(* IEC 61131-3 sources: volt/packages/volt-lsp-iec/test-corpus/awa-palletizer/Device/Plc Logic/Application/Library Manager/L_IE1P_ApplicationErrorsImplementation, 41 files *)

(* ---- L_IE1P_ERRORINFO.dut ---- *)
TYPE L_IE1P_ERRORINFO :
STRUCT
	XERROR : BOOL;
	WTEXTREFID : WORD;
	WERRORID : WORD;
	ESEVERITY : L_IE1P_SeverityLevel;
	EREACTION : L_IE1P_Reaction;
	EGROUP : L_IE1P_Group;
END_STRUCT
END_TYPE

(* ---- L_IE1P_ERRORINFORMATION.dut ---- *)
TYPE L_IE1P_ERRORINFORMATION :
STRUCT
	EERRORID : L_IE1P_Error;
	WCOMPID : WORD;
	ESEVERITY : L_IE1P_SeverityLevel;
	PSINSTANCENAME : POINTER TO STRING;
	INSTANCEID : DWORD := 0;
	TTIMESTAMP : TIME;
	TRESETTIMESTAMP : TIME;
	XCYCLIC : BOOL;
	DWEXTENDEDERRORINFO : DWORD;
	XEXTERNALERROR : BOOL;
	XCLEARERRORNEEDED : BOOL;
END_STRUCT
END_TYPE

(* ---- L_IE1P_INSTANCEIDS.dut ---- *)
TYPE L_IE1P_INSTANCEIDS :
STRUCT
	EXTINSTANCEID : DWORD;
	ADDINSTANCID1 : DWORD;
	ADDINSTANCID2 : DWORD;
	ADDINSTANCID3 : DWORD;
	ADDINSTANCID4 : DWORD;
END_STRUCT
END_TYPE

(* ---- L_IE1P_PARAMETERITEMMID.dut ---- *)
TYPE L_IE1P_PARAMETERITEMMID :
STRUCT
	SIZE : BYTE;
	ETYPE : INT;
	VALUE : L_IE1P_ParaValueMid;
END_STRUCT
END_TYPE

(* ---- L_IE1P_PARAVALUEMID.dut ---- *)
TYPE L_IE1P_PARAVALUEMID :
UNION
	DWVALUE : DWORD;
	DIVALUE : DINT;
	LRVALUE : REAL;
	SVALUE : STRING;
END_UNION
END_TYPE

(* ---- L_IE1P_PLACEHOLDERTYPE.dut ---- *)
TYPE L_IE1P_PLACEHOLDERTYPE :
(
	VTNONE := 0,
	VTDINT := 4,
	VTDWORD := 7,
	VTSTRING := 9
);
END_TYPE

(* ---- L_IE1P_PLACEHOLDERVALUE.dut ---- *)
TYPE L_IE1P_PLACEHOLDERVALUE :
UNION
	DIVALUE : DINT;
	DWVALUE : DWORD;
	RVALUE : REAL;
	LRVALUE : LREAL;
	SVALUE : STRING(50);
END_UNION
END_TYPE

(* ---- L_IE1P_PLACEHOLDERVARIABLE.dut ---- *)
TYPE L_IE1P_PLACEHOLDERVARIABLE :
STRUCT
	VARTYPE : L_IE1P_PlaceHolderType;
	VALUE : L_IE1P_PlaceholderValue;
END_STRUCT
END_TYPE

(* ---- L_IE1P_INTERNAL.gvl ---- *)
VAR_GLOBAL
	DEVICEEVENTMONITOR : L_IE1P_DeviceEventMonitor;
END_VAR

(* ---- L_IE1P_IATTRIBUTES.itf ---- *)
INTERFACE L_IE1P_IATTRIBUTES
END_INTERFACE

METHOD GET1STATTRIBUTE : DINT
END_METHOD

METHOD GET2NDATTRIBUTE : LREAL
END_METHOD

METHOD GET3RDATTRIBUTE : STRING(20)
END_METHOD

(* ---- L_IE1P_ITEXTPLACEHOLDER.itf ---- *)
INTERFACE L_IE1P_ITEXTPLACEHOLDER
END_INTERFACE

METHOD GETPLACEHOLDERDATA : L_IE1P_PlaceHolderType
VAR_INPUT
	INDEX : WORD;
END_VAR
VAR_OUTPUT
	PDATA : POINTER TO BYTE;
END_VAR
END_METHOD

(* ---- GETBOOLEANPROPERTY.pou ---- *)
FUNCTION GETBOOLEANPROPERTY : BOOL
VAR_INPUT
	STKEY : WSTRING;
END_VAR
END_FUNCTION

(* ---- GETCOMPANY.pou ---- *)
FUNCTION GETCOMPANY : WSTRING
END_FUNCTION

(* ---- GETNUMBERPROPERTY.pou ---- *)
FUNCTION GETNUMBERPROPERTY : DINT
VAR_INPUT
	STKEY : WSTRING;
END_VAR
END_FUNCTION

(* ---- GETTEXTPROPERTY.pou ---- *)
FUNCTION GETTEXTPROPERTY : WSTRING
VAR_INPUT
	STKEY : WSTRING;
END_VAR
END_FUNCTION

(* ---- GETTEXTPROPERTY2.pou ---- *)
FUNCTION GETTEXTPROPERTY2 : POINTER TO WSTRING
VAR_INPUT
	STKEY : WSTRING;
END_VAR
END_FUNCTION

(* ---- GETTITLE.pou ---- *)
FUNCTION GETTITLE : WSTRING
END_FUNCTION

(* ---- GETVERSION.pou ---- *)
FUNCTION GETVERSION : VERSION
END_FUNCTION

(* ---- GETVERSIONPROPERTY.pou ---- *)
FUNCTION GETVERSIONPROPERTY : VERSION
VAR_INPUT
	STKEY : WSTRING;
END_VAR
END_FUNCTION

(* ---- L_IE1P_GETHIGHESTREACTION.pou ---- *)
FUNCTION L_IE1P_GETHIGHESTREACTION : BOOL
VAR_INPUT
	EREACTION1 : L_IE1P_Reaction;
	MODULEHANDLER1 : POINTER TO BYTE;
	EREACTION2 : L_IE1P_Reaction;
	MODULEHANDLER2 : POINTER TO BYTE;
END_VAR
VAR_OUTPUT
	EREACTION : L_IE1P_Reaction;
	MODULEHANDLER : POINTER TO BYTE;
END_VAR
END_FUNCTION

(* ---- L_IE1P_GETHIGHESTSEVERITYANDREACTION.pou ---- *)
FUNCTION L_IE1P_GETHIGHESTSEVERITYANDREACTION : BOOL
VAR_INPUT
	ESEVERITY1 : L_IE1P_SeverityLevel;
	EREACTION1 : L_IE1P_Reaction;
	MODULEHANDLER1 : POINTER TO BYTE;
	ESEVERITY2 : L_IE1P_SeverityLevel;
	EREACTION2 : L_IE1P_Reaction;
	MODULEHANDLER2 : POINTER TO BYTE;
END_VAR
VAR_OUTPUT
	ESEVERITY : L_IE1P_SeverityLevel;
	EREACTION : L_IE1P_Reaction;
	MODULEHANDLER : POINTER TO BYTE;
END_VAR
END_FUNCTION

(* ---- L_IE1P_READERRORDATAFROMCOMPONENTLIST.pou ---- *)
FUNCTION L_IE1P_READERRORDATAFROMCOMPONENTLIST : BOOL
VAR_INPUT
	MODULEHANDLE : UDINT;
	PDATA : POINTER TO L_IE1P_ReadErrorData;
END_VAR
VAR_OUTPUT
	SEVERITY : L_IE1P_SeverityLevel;
	ERRORCODE : DWORD := 0;
END_VAR
VAR_IN_OUT
	DWCOMPIDX : DWORD;
END_VAR
END_FUNCTION

(* ---- GLOBALTEXTLIST.pou ---- *)
FUNCTION_BLOCK GLOBALTEXTLIST
VAR
	M_TEXTLISTFILE : STRING(255);
	_STNAMESPACE : STRING;
END_VAR
END_FUNCTION_BLOCK

(* ---- L_IE1P_ATTRIBUTES.pou ---- *)
FUNCTION_BLOCK L_IE1P_ATTRIBUTES
VAR_INPUT
	DIATTRIBUTE1 : DINT;
	LRATTRIBUTE2 : LREAL;
	SATTRIBUTE3 : STRING(20);
END_VAR
END_FUNCTION_BLOCK

METHOD GET1STATTRIBUTE : DINT
END_METHOD

METHOD GET2NDATTRIBUTE : LREAL
END_METHOD

METHOD GET3RDATTRIBUTE : STRING(20)
END_METHOD

(* ---- L_IE1P_DEVICEEVENTMONITOR.pou ---- *)
FUNCTION_BLOCK L_IE1P_DEVICEEVENTMONITOR
VAR
	ITFCALLBACK : CmpEventMgr.ICmpEventCallback;
	HEVENTACTUALERROR : SysTypes.RTS_IEC_HANDLE := SysTypes.RTS_INVALID_HANDLE;
	HINTERFACEACTUALERROR : SysTypes.RTS_IEC_HANDLE := SysTypes.RTS_INVALID_HANDLE;
	DWERRORUPDATED : DWORD := 0;
	AEACTSEVERITY : ARRAY [1..2] OF L_IE1P_SeverityLevel;
	ADWACTERRORCODE : ARRAY [1..2] OF DWORD;
	USIACTIVEERRORINFO : USINT;
END_VAR
END_FUNCTION_BLOCK

METHOD READACTUALERRORCODE
VAR_OUTPUT
	ESEVERITY : USINT;
	EREACTION : WORD;
	DWERRORCODE : DWORD;
END_VAR
END_METHOD

METHOD EVENTCALLBACK : UDINT
VAR_INPUT
	PEVENTPARAM : POINTER TO EventParam;
END_VAR
END_METHOD

METHOD REGISTEREVENT
VAR_INPUT
	XONLYCALLBACKFUNCTION : BOOL;
END_VAR
END_METHOD

METHOD UNREGISTEREVENT
VAR_INPUT
	XONLYCALLBACKFUNCTION : BOOL;
END_VAR
END_METHOD

METHOD FB_REINIT : BOOL
END_METHOD

METHOD FB_EXIT : BOOL
VAR_INPUT
	BINCOPYCODE : BOOL;
END_VAR
END_METHOD

METHOD FB_INIT : BOOL
VAR_INPUT
	BINITRETAINS : BOOL;
	BINCOPYCODE : BOOL;
END_VAR
END_METHOD

(* ---- L_IE1P_EMPTYERRORHANDLER.pou ---- *)
FUNCTION_BLOCK L_IE1P_EMPTYERRORHANDLER
END_FUNCTION_BLOCK

METHOD ITFCHECKERRORRESETOCCURED : BOOL
VAR_IN_OUT
	RESETTIME : SYSTIME;
END_VAR
END_METHOD

METHOD ITFCLEARERROR : DWORD
VAR_INPUT
	ESEVERITY : L_IE1P_SeverityLevel;
	WERRORID : WORD;
	WCOMPID : WORD;
	DWINSTANCEID : DWORD := 0;
END_VAR
END_METHOD

METHOD ITFCLEARREACTION
VAR_INPUT
	EREACTION : L_IE1P_Reaction;
	DICLEARCOUNT : DINT;
	DWINSTANCEID : DWORD;
END_VAR
END_METHOD

METHOD ITFGETACTUALERRORCODE : DWORD
VAR_OUTPUT
	ESEVERITY : WORD;
END_VAR
END_METHOD

METHOD ITFREGISTERERRORINSTANCE : DWORD
END_METHOD

METHOD ITFRESETACTIVE : BOOL
END_METHOD

METHOD ITFRESETERROR : DWORD
VAR_INPUT
	ERRORHANDLE : RTS_IEC_HANDLE := 0;
END_VAR
END_METHOD

METHOD ITFRESETERRORREACTION
VAR_INPUT
	DWINSTANCEID : DWORD := 0;
END_VAR
END_METHOD

METHOD ITFSETERROR : DWORD
VAR_INPUT
	ESEVERITY : L_IE1P_SeverityLevel;
	WERRORID : WORD;
	WCOMPID : WORD;
	DWINSTANCEID : DWORD := 0;
	EREACTION : L_IE1P_Reaction;
END_VAR
END_METHOD

(* ---- L_IE1P_ERRORHANDLER.pou ---- *)
FUNCTION_BLOCK L_IE1P_ERRORHANDLER
VAR_INPUT
	ADDERRORHANDLER1 : L_IE1P_IErrorHandler;
	ADDERRORHANDLER2 : L_IE1P_IErrorHandler;
	ADDERRORHANDLER3 : L_IE1P_IErrorHandler;
	ADDERRORHANDLER4 : L_IE1P_IErrorHandler;
END_VAR
VAR_OUTPUT
	XWARNINGACTIVE : BOOL;
	XWARNINGLOCKACTIVE : BOOL;
	XFAULTQSPAPPLACTIVE : BOOL;
	XFAULTQSPACTIVE : BOOL;
	XFAULTQSPCINHACTIVE : BOOL;
	XFAULTACTIVE : BOOL;
END_VAR
VAR
	ERRORMANAGER : L_IE1P_ErrorManager;
	ADDERRORHANDLERINSTANCEIDS : ARRAY [1..MaxInstanceIDs] OF L_IE1P_InstanceIDs;
	ERRORRESETOCCUREDTIME : SysTime;
	C_STRUNDEFERROR : STRING := 'undefined';
	MAXINSTANCEIDS : WORD := 15;
END_VAR
END_FUNCTION_BLOCK

METHOD CHECKHIGHESTSEVERITY
VAR_INPUT
	ESEVERITYNEW : WORD;
	DWERRORCODENEW : DWORD;
END_VAR
VAR_IN_OUT
	ESEVERITYACT : WORD;
	DWERRORCODEACT : DWORD;
END_VAR
END_METHOD

METHOD FINDADDINSTANCEID : DWORD
VAR_INPUT
	DWEXTINSTANCEID : DWORD;
	DWNUMBER : DWORD;
END_VAR
END_METHOD

METHOD FB_INIT : BOOL
VAR_INPUT
	BINITRETAINS : BOOL;
	BINCOPYCODE : BOOL;
END_VAR
END_METHOD

METHOD ITFCHECKERRORRESETOCCURED : BOOL
VAR_IN_OUT
	RESETTIME : SYSTIME;
END_VAR
END_METHOD

METHOD ITFCLEARERROR : DWORD
VAR_INPUT
	ESEVERITY : L_IE1P_SeverityLevel;
	WERRORID : WORD;
	WCOMPID : WORD;
	DWINSTANCEID : DWORD := 0;
END_VAR
END_METHOD

METHOD ITFCLEARREACTION
VAR_INPUT
	EREACTION : L_IE1P_Reaction;
	DICLEARCOUNT : DINT;
	DWINSTANCEID : DWORD;
END_VAR
END_METHOD

METHOD ITFGETACTUALERRORCODE : DWORD
VAR_OUTPUT
	ESEVERITY : WORD;
END_VAR
END_METHOD

METHOD ITFREGISTERERRORINSTANCE : DWORD
END_METHOD

METHOD ITFRESETACTIVE : BOOL
END_METHOD

METHOD ITFRESETERROR : DWORD
VAR_INPUT
	ERRORHANDLE : RTS_IEC_HANDLE := 0;
END_VAR
END_METHOD

METHOD ITFRESETERRORREACTION
VAR_INPUT
	DWINSTANCEID : DWORD := 0;
END_VAR
END_METHOD

METHOD ITFSETERROR : DWORD
VAR_INPUT
	ESEVERITY : L_IE1P_SeverityLevel;
	WERRORID : WORD;
	WCOMPID : WORD;
	DWINSTANCEID : DWORD := 0;
	EREACTION : L_IE1P_Reaction;
END_VAR
END_METHOD

(* ---- L_IE1P_ERRORMANAGER.pou ---- *)
FUNCTION_BLOCK L_IE1P_ERRORMANAGER
VAR_INPUT
	XUSEADDLOGIPC : BOOL := TRUE;
	DWTASKYCLE_US : DWORD := 1000;
	XIGNOREFAULT_LOG : BOOL := TRUE;
	XNOLOGBOOKENTRY : BOOL := FALSE;
END_VAR
VAR
	EACTIVEERRORID : REFERENCE TO L_IE1P_Error;
	EACTIVESEVERITY : REFERENCE TO L_IE1P_SeverityLevel;
	XERROR : REFERENCE TO BOOL;
	XWARNING : REFERENCE TO BOOL;
	PSERRORINST : REFERENCE TO POINTER TO STRING;
	SERRORINST : REFERENCE TO STRING;
	IACTIVEERRORENTRY : INT;
	IACTIVEWARNINGENTRY : INT;
	IFIRSTERROR : INT;
	IFIRSTWARNING : INT;
	PSERRORINSTOLD : POINTER TO STRING;
	DWERRORITFID : DWORD := 0;
	ASCERRORINFO : ARRAY [0..7] OF L_IE1P_ErrorInformation;
	ASCWARNINGINFO : ARRAY [0..7] OF L_IE1P_ErrorInformation;
	MODULEHANDLER_INT : L_IMHP_IModuleHandler;
	DUMMY_EACTIVEERRORID : L_IE1P_Error;
	DUMMY_EACTIVESEVERITY : L_IE1P_SeverityLevel;
	DUMMY_XERROR : BOOL;
	DUMMY_XWARNING : BOOL;
	DUMMY_PSERRORINST : POINTER TO STRING;
	DUMMY_SERRORINST : STRING;
	C_STRNOERROR : STRING := '-';
	C_STRUNDEFERROR : STRING := 'undefined';
END_VAR
END_FUNCTION_BLOCK

METHOD ADDERRORENTRY : BOOL
VAR_INPUT
	WERRORID : L_IE1P_Error := 0;
	WCOMPID : WORD;
	ESEVERITY : L_IE1P_SeverityLevel;
	INSTANCEID : DWORD := 0;
	PSINSTANCENAME : POINTER TO BYTE := 0;
	DWEXTENDEDERRORINFO : DWORD;
	XAUTORESET : BOOL;
	XEXTERNALERROR : BOOL;
END_VAR
VAR_OUTPUT
	PERRORINFO : POINTER TO L_IE1P_ErrorInformation;
END_VAR
END_METHOD

METHOD CLEARERRORENTRY
VAR_INPUT
	INSTANCEID : DWORD := 0;
	WERRORID : WORD;
	DWEXTENDEDERRORINFO : DWORD;
END_VAR
END_METHOD

METHOD COUNTEXTERNALERROR : INT
VAR_OUTPUT
	OTHERERRORS : INT := 0;
END_VAR
END_METHOD

METHOD CYCLICUPDATEERRORINFO
END_METHOD

METHOD ERRORRESETPOSSIBLE : BOOL
VAR_OUTPUT
	EACTSEVERITY : L_IE1P_SeverityLevel;
END_VAR
END_METHOD

METHOD ERRORRESETPOSSIBLEWITHOUTEXTERNAL : BOOL
VAR_OUTPUT
	EACTSEVERITY : L_IE1P_SeverityLevel;
END_VAR
END_METHOD

METHOD FINDANDDELETEERRORENTRY : BOOL
VAR_INPUT
	DWINSTANCEID : DWORD := 0;
	XEXTERNAL : BOOL;
	XEXTERNALERRORRESETHANDLING : BOOL := FALSE;
END_VAR
END_METHOD

METHOD GENLOGENTRY
VAR_INPUT
	ERRORHANDLE : SysTypes.RTS_IEC_HANDLE;
	WERRORID : L_IE1P_Error := L_IE1P_Error.NoError;
	WCOMPID : WORD;
	ESEVERITY : L_IE1P_SeverityLevel;
	DWEXTENDEDERRORINFO : DWORD;
	INSTANCEID : DWORD := 0;
	PSINSTANCENAME : POINTER TO BYTE := 0;
	PERRORINFO : POINTER TO L_IE1P_ErrorInformation := 0;
END_VAR
END_METHOD

METHOD GETERRORITFID : DWORD
END_METHOD

METHOD INITIALIZE
VAR_INPUT
	PEACTIVEERRORID : POINTER TO L_IE1P_Error;
	PXERROR : POINTER TO BOOL;
	PXWARNING : POINTER TO BOOL;
	PPSERRORINST : POINTER TO POINTER TO STRING;
	PSERRORINST : POINTER TO STRING;
END_VAR
END_METHOD

METHOD RESET
END_METHOD

METHOD RESETERRORDATA
VAR_IN_OUT
	ERRORINFO : L_IE1P_ErrorInformation;
END_VAR
END_METHOD

METHOD RESETERRORINFO
END_METHOD

METHOD RESETWARNINGINFO
END_METHOD

METHOD SETMODULEHANDLER : BOOL
VAR_INPUT
	MODULEHANDLER : L_IMHP_IModuleHandler;
END_VAR
END_METHOD

METHOD UPDATEERRORINFO
END_METHOD

METHOD FB_INIT : BOOL
VAR_INPUT
	BINITRETAINS : BOOL;
	BINCOPYCODE : BOOL;
END_VAR
END_METHOD

(* ---- L_IE1P_FORWARDERROR.pou ---- *)
FUNCTION_BLOCK L_IE1P_FORWARDERROR
VAR_INPUT
	XENABLE : BOOL;
	MODULEHANDLER : L_IMHP_IModuleHandler;
	XRESETERROR : BOOL;
	XERRORACTIVE : BOOL;
	XWARNINGACTIVE : BOOL;
	WERRORID : WORD;
	WTEXTREFID : WORD;
	ERRORMODULEHANDLER : L_IMHP_IModuleHandler;
END_VAR
VAR_OUTPUT
	XBUSY : BOOL;
	XERROR : BOOL;
	EERRORID : L_IE1P_Error;
	XERRORRESETACTIVE : BOOL;
END_VAR
VAR
	ERRORHANDLE : SysTypes.RTS_IEC_HANDLE;
	XERROROLD : BOOL;
	XWARNINGOLD : BOOL;
	WERRORIDOLD : WORD;
	WTEXTREFIDOLD : WORD;
	XENABLEOLD : BOOL;
	ITFCALLBACK : CmpEventMgr.ICmpEventCallback;
	HEVENTRESETOCCURED : SysTypes.RTS_IEC_HANDLE := SysTypes.RTS_INVALID_HANDLE;
	HINTERFACERESETOCCURED : SysTypes.RTS_IEC_HANDLE := SysTypes.RTS_INVALID_HANDLE;
	WEVTCOUNT_RESETOCCURED : WORD;
	XRESETOCCURED : BOOL;
	XRESETERROROLD : BOOL;
	LRCYCLESERRORRESETACTIVE : LREAL;
	XERRORRESETACTIVEINTERN : BOOL;
	WRESETCOUNTER : WORD;
	WRESETSUSPENDCOUNTER : WORD;
	XWARNINGSEVACTIVE : BOOL;
	XERRORSEVACTIVE : BOOL;
	XWARNINGTEXTREFID : BOOL;
	XERRORTEXTREFID : BOOL;
	C_WARNING : USINT := 2;
	C_ERROR : USINT := 18;
	WARNING_TEXTREFID : WORD := L_IE1P_Error.DriveWarningMsgNotResolvable;
	ERROR_TEXTREFID : WORD := L_IE1P_Error.DriveErrorMsgNotResolvable;
	INTERNALERRORTEXTREFID : WORD := 16#2C00;
	DEFAULT_TEXTREFID : WORD := 16#2009;
END_VAR
END_FUNCTION_BLOCK

METHOD FB_REINIT : BOOL
END_METHOD

METHOD FB_EXIT : BOOL
VAR_INPUT
	BINCOPYCODE : BOOL;
END_VAR
END_METHOD

METHOD FB_INIT : BOOL
VAR_INPUT
	BINITRETAINS : BOOL;
	BINCOPYCODE : BOOL;
END_VAR
END_METHOD

METHOD EVENTCALLBACK : UDINT
VAR_INPUT
	PEVENTPARAM : POINTER TO EventParam;
END_VAR
END_METHOD

METHOD REGISTEREVENT
VAR_INPUT
	XONLYCALLBACKFUNCTION : BOOL;
END_VAR
END_METHOD

METHOD UNREGISTEREVENT
VAR_INPUT
	XONLYCALLBACKFUNCTION : BOOL;
END_VAR
END_METHOD

(* ---- L_IE1P_FORWARDSEVERITY.pou ---- *)
FUNCTION_BLOCK L_IE1P_FORWARDSEVERITY
VAR_INPUT
	XENABLE : BOOL;
	MODULEHANDLER : L_IMHP_IModuleHandler;
	XFORWARDFROMCHILDMODULES : BOOL;
	XDISABLEFORWARDTOPARENT : BOOL;
END_VAR
VAR_OUTPUT
	XBUSY : BOOL;
	XERROR : BOOL;
	EERRORID : L_IE1P_Error;
END_VAR
VAR
	XENABLEOLD : BOOL;
	XFORWARDSEVERITYSUBMODULESCALLED : BOOL;
END_VAR
END_FUNCTION_BLOCK

(* ---- L_IE1P_READACTUALERRORCODE.pou ---- *)
FUNCTION_BLOCK L_IE1P_READACTUALERRORCODE
VAR_INPUT
	XENABLE : BOOL;
	MODULEHANDLER : L_IMHP_IModuleHandler;
	ERRORHANDLER : L_IE1P_IErrorHandler;
END_VAR
VAR_OUTPUT
	XBUSY : BOOL;
	XERROR : BOOL;
	EERRORID : L_IE1P_Error;
	XERRORACTIVE : BOOL;
	XWARNINGACTIVE : BOOL;
	DWERRORCODE : DWORD;
	ESEVERITY : L_IE1P_SeverityLevel;
END_VAR
VAR
	SEVTMP : WORD;
	XACTUALERRORFROMMODULESUPPORTED : BOOL := FALSE;
	MYMODULETMP : L_IMHP_IModuleHandler;
	EREACTIONTMP : L_IE1P_Reaction;
END_VAR
END_FUNCTION_BLOCK

METHOD FB_EXIT : BOOL
VAR_INPUT
	BINCOPYCODE : BOOL;
END_VAR
END_METHOD

METHOD FB_INIT : BOOL
VAR_INPUT
	BINITRETAINS : BOOL;
	BINCOPYCODE : BOOL;
END_VAR
END_METHOD

(* ---- L_IE1P_READACTUALSEVERITY.pou ---- *)
FUNCTION_BLOCK L_IE1P_READACTUALSEVERITY
VAR_INPUT
	XENABLE : BOOL;
	MODULEHANDLER : L_IMHP_IModuleHandler;
	XDISABLESUBMODULES : BOOL;
	XINCLUDEOWNMODULE : BOOL := TRUE;
	XONLYSUBMODULES : BOOL := FALSE;
END_VAR
VAR_OUTPUT
	XBUSY : BOOL;
	XERROR : BOOL;
	EERRORID : L_IE1P_Error;
	ESEVERITY : L_IE1P_SeverityLevel;
	EREACTION : L_IE1P_Reaction;
	SAFFECTEDMODULENAME : STRING;
	AFFECTEDMODULEHANDLER : L_IMHP_IModuleHandler;
	XERRORACTIVE : BOOL;
	XWARNINGACTIVE : BOOL;
	SEVERITYSTATUS : L_IE1P_SeverityStatus;
	REACTIONSTATUS : L_IE1P_ReactionStatus;
END_VAR
VAR
	XENABLEOLD : BOOL;
	AFFECTEDMODULEHANDLEROLD : L_IMHP_IModuleHandler;
	MODULEHANDLER_INT : L_IMHP_IModuleHandler;
	XDUMMY : BOOL;
END_VAR
END_FUNCTION_BLOCK

METHOD READCHILDSEVERITY : BOOL
VAR_INPUT
	WCHILD : WORD;
END_VAR
VAR_OUTPUT
	ESEVERITY : L_IE1P_SeverityLevel;
	EREACTION : L_IE1P_Reaction;
	SCHILDNAME : STRING;
	CHILDMODULEHANDER : L_IMHP_IModuleHandler;
END_VAR
END_METHOD

(* ---- L_IE1P_READCURRENTERROR.pou ---- *)
FUNCTION_BLOCK L_IE1P_READCURRENTERROR
VAR_INPUT
	XENABLE : BOOL;
END_VAR
VAR_OUTPUT
	XBUSY : BOOL;
	XERROR : BOOL;
	EERRORID : L_IE1P_Error;
	XERRORACTIVE : BOOL;
	XWARNINGACTIVE : BOOL;
	DWERRORCODE : DWORD;
	ESEVERITY : L_IE1P_SeverityLevel;
END_VAR
VAR
	XENABLEOLD : BOOL;
	EREACTIONTMP : L_IE1P_Reaction;
END_VAR
END_FUNCTION_BLOCK

(* ---- L_IE1P_RESETERROR.pou ---- *)
FUNCTION_BLOCK L_IE1P_RESETERROR
VAR_INPUT
	MODULEHANDLER : L_IMHP_IModuleHandler;
	ERRORHANDLER : L_IE1P_IErrorHandler;
	XRESETERROR : BOOL;
END_VAR
VAR_OUTPUT
	XERROR : BOOL;
	EERRORID : L_IE1P_Error;
	XERRORRESETACTIVE : BOOL;
	XRESETACTIVE : BOOL;
END_VAR
VAR
	MODULEHANDLER_INT : L_IMHP_IModuleHandler := 0;
	EXTMODULEHANDLER : L_IMHP_IModuleHandler := 0;
	ERRORHANDLE : SysTypes.RTS_IEC_HANDLE := 0;
	ITFCALLBACK : CmpEventMgr.ICmpEventCallback;
	HEVENTRESETOCCURED : SysTypes.RTS_IEC_HANDLE := SysTypes.RTS_INVALID_HANDLE;
	HINTERFACERESETOCCURED : SysTypes.RTS_IEC_HANDLE := SysTypes.RTS_INVALID_HANDLE;
	WEVTCOUNT_RESETOCCURED : WORD;
	XRESETOCCURED : BOOL;
	XRESETERROROLD : BOOL;
	XRESETERROROLD2 : BOOL;
	ERRORRESETTRIGGERTIME : TIME;
END_VAR
END_FUNCTION_BLOCK

METHOD FB_REINIT : BOOL
END_METHOD

METHOD RESETERRORCOMPLIST
END_METHOD

METHOD FB_EXIT : BOOL
VAR_INPUT
	BINCOPYCODE : BOOL;
END_VAR
END_METHOD

METHOD FB_INIT : BOOL
VAR_INPUT
	BINITRETAINS : BOOL;
	BINCOPYCODE : BOOL;
END_VAR
END_METHOD

METHOD EVENTCALLBACK : UDINT
VAR_INPUT
	PEVENTPARAM : POINTER TO EventParam;
END_VAR
END_METHOD

METHOD REGISTEREVENT
VAR_INPUT
	XONLYCALLBACKFUNCTION : BOOL;
END_VAR
END_METHOD

METHOD UNREGISTEREVENT
VAR_INPUT
	XONLYCALLBACKFUNCTION : BOOL;
END_VAR
END_METHOD

(* ---- L_IE1P_RESETERRORGLOBAL.pou ---- *)
FUNCTION_BLOCK L_IE1P_RESETERRORGLOBAL
VAR_INPUT
	XRESETERROR : BOOL;
END_VAR
VAR_OUTPUT
	XERROR : BOOL;
	EERRORID : L_IE1P_Error;
	XERRORRESETACTIVE : BOOL;
END_VAR
VAR
	EXTMODULEHANDLER : L_IMHP_IModuleHandler := 0;
	ERRORHANDLE : SysTypes.RTS_IEC_HANDLE := 0;
	ITFCALLBACK : CmpEventMgr.ICmpEventCallback;
	HEVENTRESETOCCURED : SysTypes.RTS_IEC_HANDLE := SysTypes.RTS_INVALID_HANDLE;
	HINTERFACERESETOCCURED : SysTypes.RTS_IEC_HANDLE := SysTypes.RTS_INVALID_HANDLE;
	WEVTCOUNT_RESETOCCURED : WORD;
	XRESETOCCURED : BOOL;
	XRESETERROROLD : BOOL;
END_VAR
END_FUNCTION_BLOCK

METHOD FB_REINIT : BOOL
END_METHOD

METHOD FB_EXIT : BOOL
VAR_INPUT
	BINCOPYCODE : BOOL;
END_VAR
END_METHOD

METHOD FB_INIT : BOOL
VAR_INPUT
	BINITRETAINS : BOOL;
	BINCOPYCODE : BOOL;
END_VAR
END_METHOD

METHOD EVENTCALLBACK : UDINT
VAR_INPUT
	PEVENTPARAM : POINTER TO EventParam;
END_VAR
END_METHOD

METHOD REGISTEREVENT
VAR_INPUT
	XONLYCALLBACKFUNCTION : BOOL;
END_VAR
END_METHOD

METHOD UNREGISTEREVENT
VAR_INPUT
	XONLYCALLBACKFUNCTION : BOOL;
END_VAR
END_METHOD

(* ---- L_IE1P_SETERROR.pou ---- *)
FUNCTION_BLOCK L_IE1P_SETERROR
VAR_INPUT
	MODULEHANDLER : L_IMHP_IModuleHandler;
	ERRORHANDLER : L_IE1P_IErrorHandler;
	WTEXTREFID : WORD;
	XRESETERROR : BOOL;
	XSETERROR1 : BOOL;
	ESEVERITY1 : L_IE1P_SeverityLevel;
	WERRORID1 : WORD;
	WTEXTREFID1 : WORD;
	EREACTION1 : L_IE1P_Reaction := L_IE1P_Reaction.No_Reaction;
	EGROUP1 : L_IE1P_Group := L_IE1P_Group.ManufacturerGroup;
	XSETERROR2 : BOOL;
	ESEVERITY2 : L_IE1P_SeverityLevel;
	WERRORID2 : WORD;
	WTEXTREFID2 : WORD;
	EREACTION2 : L_IE1P_Reaction := L_IE1P_Reaction.No_Reaction;
	EGROUP2 : L_IE1P_Group := L_IE1P_Group.ManufacturerGroup;
	XSETERROR3 : BOOL;
	ESEVERITY3 : L_IE1P_SeverityLevel;
	WERRORID3 : WORD;
	WTEXTREFID3 : WORD;
	EREACTION3 : L_IE1P_Reaction := L_IE1P_Reaction.No_Reaction;
	EGROUP3 : L_IE1P_Group := L_IE1P_Group.ManufacturerGroup;
	XSETERROR4 : BOOL;
	ESEVERITY4 : L_IE1P_SeverityLevel;
	WERRORID4 : WORD;
	WTEXTREFID4 : WORD;
	EREACTION4 : L_IE1P_Reaction := L_IE1P_Reaction.No_Reaction;
	EGROUP4 : L_IE1P_Group := L_IE1P_Group.ManufacturerGroup;
END_VAR
VAR_OUTPUT
	XERROR : BOOL;
	EERRORID : L_IE1P_Error;
	XERRORRESETACTIVE : BOOL;
	SCERRORINFORMATION1 : L_IE1P_ErrorInfo;
	SCERRORINFORMATION2 : L_IE1P_ErrorInfo;
	SCERRORINFORMATION3 : L_IE1P_ErrorInfo;
	SCERRORINFORMATION4 : L_IE1P_ErrorInfo;
END_VAR
VAR
	XREGISTEROVERSEMP : BOOL := FALSE;
	XRESETERROROLD : BOOL;
	XSETERROR1OLD : BOOL;
	XSETERROR2OLD : BOOL;
	XSETERROR3OLD : BOOL;
	XSETERROR4OLD : BOOL;
	ESEVERITY1_INT : L_IE1P_SeverityLevel;
	ESEVERITY2_INT : L_IE1P_SeverityLevel;
	ESEVERITY3_INT : L_IE1P_SeverityLevel;
	ESEVERITY4_INT : L_IE1P_SeverityLevel;
	WTEXTREFID1_INT : WORD;
	WTEXTREFID2_INT : WORD;
	WTEXTREFID3_INT : WORD;
	WTEXTREFID4_INT : WORD;
	WERRORID1_INT : WORD;
	WERRORID2_INT : WORD;
	WERRORID3_INT : WORD;
	WERRORID4_INT : WORD;
	EREACTION1_INT : L_IE1P_Reaction;
	EREACTION2_INT : L_IE1P_Reaction;
	EREACTION3_INT : L_IE1P_Reaction;
	EREACTION4_INT : L_IE1P_Reaction;
	XFBERRORINT1 : BOOL;
	EFBERRORIDINT1 : L_IE1P_Error;
	XFBERRORINT2 : BOOL;
	EFBERRORIDINT2 : L_IE1P_Error;
	XFBERRORINT3 : BOOL;
	EFBERRORIDINT3 : L_IE1P_Error;
	XFBERRORINT4 : BOOL;
	EFBERRORIDINT4 : L_IE1P_Error;
	ERRORHANDLEINTERNAL : SysTypes.RTS_IEC_HANDLE := 0;
	ERRORHANDLEACT : SysTypes.RTS_IEC_HANDLE := 0;
	ERRORHANDLEINT1 : SysTypes.RTS_IEC_HANDLE := 0;
	ERRORHANDLEINT2 : SysTypes.RTS_IEC_HANDLE := 0;
	ERRORHANDLEINT3 : SysTypes.RTS_IEC_HANDLE := 0;
	ERRORHANDLEINT4 : SysTypes.RTS_IEC_HANDLE := 0;
	ITFCALLBACK : CmpEventMgr.ICmpEventCallback;
	HEVENTRESETOCCURED : SysTypes.RTS_IEC_HANDLE := SysTypes.RTS_INVALID_HANDLE;
	HINTERFACERESETOCCURED : SysTypes.RTS_IEC_HANDLE := SysTypes.RTS_INVALID_HANDLE;
	WEVTCOUNT_RESETOCCURED : WORD;
	XRESETOCCURED : BOOL;
	XFIRSTCYCLE : BOOL := FALSE;
	DWINSTANCEID : DWORD;
	REACTIONCOUNTERINFORMATIONNOTIFY : L_IE1P_ReactionCounter;
	REACTIONCOUNTERINFORMATIONCLEAR : L_IE1P_ReactionCounter;
	REACTIONCOUNTERWARNINGNOTIFY : L_IE1P_ReactionCounter;
	REACTIONCOUNTERWARNINGCLEAR : L_IE1P_ReactionCounter;
	REACTIONCOUNTERWARNINGLOCKNOTIFY : L_IE1P_ReactionCounter;
	REACTIONCOUNTERWARNINGLOCKCLEAR : L_IE1P_ReactionCounter;
	REACTIONCOUNTERFAULTLOGNOTIFY : L_IE1P_ReactionCounter;
	REACTIONCOUNTERFAULTLOGCLEAR : L_IE1P_ReactionCounter;
	REACTIONCOUNTERFAULTNOTIFY : L_IE1P_ReactionCounter;
	REACTIONCOUNTERFAULTCLEAR : L_IE1P_ReactionCounter;
	SEVERITYCOUNTERNOTIFY : L_IE1P_SeverityCounter;
	SEVERITYCOUNTERCLEAR : L_IE1P_SeverityCounter;
	DUMMYERRORHANDLER : L_IE1P_EmptyErrorHandler;
	ERRORHANDLER_INT : L_IE1P_IErrorHandler;
	ERRORHANDLER_OLD : L_IE1P_IErrorHandler;
	MODULEHANDLER_INT : L_IMHP_IModuleHandler;
	MODULEHANDLER_OLD : L_IMHP_IModuleHandler;
	RESETTIMEERRORHANDLER : SYSTIME;
	SCOMPONENTNAME : STRING := '';
	SINSTANCESTR : STRING;
	SINSTANCESTRDUMMY : STRING;
	SCOMPNAME : STRING := '';
	COMPONENTNAME : STRING;
END_VAR
END_FUNCTION_BLOCK

METHOD AFTERGLOBALINIT
END_METHOD

METHOD CHECKSETERROR
VAR_IN_OUT
	XSETERROR : BOOL;
	XSETERROROLD : BOOL;
	ESEVERITY : L_IE1P_SeverityLevel;
	ESEVERITY_INT : L_IE1P_SeverityLevel;
	WERRORID : WORD;
	WERRORID_INT : WORD;
	WTEXTREFID : WORD;
	WTEXTREFID_INT : WORD;
	XFBERRORINT : BOOL;
	EFBERRORIDINT : L_IE1P_Error;
	EREACTION : L_IE1P_Reaction;
	EREACTION_INT : L_IE1P_Reaction;
	EGROUP : L_IE1P_Group;
	ERRORHANDLEUSED : SysTypes.RTS_IEC_HANDLE;
	SCERRORINFORMATION : L_IE1P_ErrorInfo;
END_VAR
END_METHOD

METHOD CLEANREACTIONCOUNT : DINT
VAR_INPUT
	ESEVERITY : L_IE1P_SeverityLevel;
END_VAR
VAR_IN_OUT
	REACTIONCOUNTERNOTIFY : L_IE1P_ReactionCounter;
	REACTIONCOUNTERCLEAR : L_IE1P_ReactionCounter;
END_VAR
END_METHOD

METHOD CLEANSEVERITYANDREACTIONCOUNTER
END_METHOD

METHOD CLEARERRORACTIVESTRUCT
END_METHOD

METHOD FB_REINIT : BOOL
END_METHOD

METHOD GETINSTANCENAME : STRING
END_METHOD

METHOD SETREACTIONCOUNTERVARIABLE
VAR_INPUT
	EREACTION : L_IE1P_Reaction;
	DICOUNT : DINT;
END_VAR
VAR_IN_OUT
	REACTIONCOUNTER : L_IE1P_ReactionCounter;
END_VAR
END_METHOD

METHOD UPDATESEVERITYANDREACTIONCOUNTER
VAR_INPUT
	WMODE : WORD;
	ESEVERITY : L_IE1P_SeverityLevel;
	EREACTION : L_IE1P_Reaction;
END_VAR
END_METHOD

METHOD FB_EXIT : BOOL
VAR_INPUT
	BINCOPYCODE : BOOL;
END_VAR
END_METHOD

METHOD FB_INIT : BOOL
VAR_INPUT
	BINITRETAINS : BOOL;
	BINCOPYCODE : BOOL;
END_VAR
END_METHOD

METHOD EVENTCALLBACK : UDINT
VAR_INPUT
	PEVENTPARAM : POINTER TO EventParam;
END_VAR
END_METHOD

METHOD REGISTEREVENT
VAR_INPUT
	XONLYCALLBACKFUNCTION : BOOL;
END_VAR
END_METHOD

METHOD UNREGISTEREVENT
VAR_INPUT
	XONLYCALLBACKFUNCTION : BOOL;
END_VAR
END_METHOD

(* ---- L_IE1P_SETERRORSINGLE.pou ---- *)
FUNCTION_BLOCK L_IE1P_SETERRORSINGLE EXTENDS L_IE1P_SetErrorSingleBase
VAR_INPUT
	MODULEHANDLER : L_IMHP_IModuleHandler;
	ERRORHANDLER : L_IE1P_IErrorHandler;
	XSETERROR : BOOL;
	ESEVERITY : L_IE1P_SeverityLevel;
	WTEXTREFID : WORD;
	WERRORID : WORD;
	EREACTION : L_IE1P_Reaction := L_IE1P_Reaction.No_Reaction;
	EGROUP : L_IE1P_Group := L_IE1P_Group.ManufacturerGroup;
	TEXTPLACEHOLDER : L_IE1P_ITextPlaceHolder;
	ATTRIBUTES : L_IE1P_IAttributes;
END_VAR
VAR_OUTPUT
	XERROR : BOOL;
	EERRORID : L_IE1P_Error;
	SCERRORINFORMATION : L_IE1P_ErrorInfo;
END_VAR
VAR
	GETCONNECTEDMODULEHANDLER : L_IMHP_IModuleHandler;
END_VAR
END_FUNCTION_BLOCK

(* ---- L_IE1P_SETERRORSINGLEBASE.pou ---- *)
FUNCTION_BLOCK L_IE1P_SETERRORSINGLEBASE
VAR
	XSETERROROLD : BOOL;
	ESEVERITY_INT : L_IE1P_SeverityLevel;
	WTEXTREFID_INT : WORD;
	WERRORID_INT : WORD;
	EREACTION_INT : L_IE1P_Reaction;
	XFBERRORINT : BOOL;
	EFBERRORIDINT : L_IE1P_Error;
	XFIRSTCYCLE : BOOL;
	ITFTEXTPLACEHOLDER_INT : L_IE1P_ITextPlaceHolder;
	ITFERRORATTRIBUTES_INT : L_IE1P_IAttributes;
	DUMMYERRORHANDLER : L_IE1P_EmptyErrorHandler;
	ERRORHANDLER_INT : L_IE1P_IErrorHandler;
	ERRORHANDLER_OLD : L_IE1P_IErrorHandler;
	MODULEHANDLER_INT : L_IMHP_IModuleHandler;
	MODULEHANDLER_OLD : L_IMHP_IModuleHandler;
	ERRORHANDLEINTERNAL : SysTypes.RTS_IEC_HANDLE := 0;
	ERRORHANDLEACT : SysTypes.RTS_IEC_HANDLE := 0;
	DWINSTANCEID : DWORD;
	ERRORHANDLEUSED : SysTypes.RTS_IEC_HANDLE := 0;
	REACTIONCOUNTERINFORMATIONNOTIFY : L_IE1P_ReactionCounter;
	REACTIONCOUNTERINFORMATIONCLEAR : L_IE1P_ReactionCounter;
	REACTIONCOUNTERWARNINGNOTIFY : L_IE1P_ReactionCounter;
	REACTIONCOUNTERWARNINGCLEAR : L_IE1P_ReactionCounter;
	REACTIONCOUNTERWARNINGLOCKNOTIFY : L_IE1P_ReactionCounter;
	REACTIONCOUNTERWARNINGLOCKCLEAR : L_IE1P_ReactionCounter;
	REACTIONCOUNTERFAULTLOGNOTIFY : L_IE1P_ReactionCounter;
	REACTIONCOUNTERFAULTLOGCLEAR : L_IE1P_ReactionCounter;
	REACTIONCOUNTERFAULTNOTIFY : L_IE1P_ReactionCounter;
	REACTIONCOUNTERFAULTCLEAR : L_IE1P_ReactionCounter;
	SEVERITYCOUNTERNOTIFY : L_IE1P_SeverityCounter;
	SEVERITYCOUNTERCLEAR : L_IE1P_SeverityCounter;
	RESETTIME : SYSTIME;
	RESETTIMEERRORHANDLER : SYSTIME;
	XRESETOCCURED : BOOL;
	XREGISTEROVERSEMP : BOOL;
	SINSTANCESTR : STRING;
	SCOMPNAME : STRING := '';
	GETCONNECTEDMODULEHANDLER : L_IMHP_IModuleHandler;
END_VAR
END_FUNCTION_BLOCK

METHOD AFTERGLOBALINIT
END_METHOD

METHOD CHECKSETERROR
VAR_IN_OUT
	XSETERROR : BOOL;
	ESEVERITY : L_IE1P_SeverityLevel;
	WERRORID : WORD;
	WTEXTREFID : WORD;
	EREACTION : L_IE1P_Reaction;
	EGROUP : L_IE1P_Group;
	SCERRORINFORMATION : L_IE1P_ErrorInfo;
END_VAR
END_METHOD

METHOD CLEANREACTIONCOUNT : DINT
VAR_INPUT
	ESEVERITY : L_IE1P_SeverityLevel;
END_VAR
VAR_IN_OUT
	REACTIONCOUNTERNOTIFY : L_IE1P_ReactionCounter;
	REACTIONCOUNTERCLEAR : L_IE1P_ReactionCounter;
END_VAR
END_METHOD

METHOD CLEANSEVERITYANDREACTIONCOUNTER
END_METHOD

METHOD GETINSTANCENAME : STRING
END_METHOD

METHOD MAIN : BOOL
VAR_IN_OUT
	MODULEHANDLER : L_IMHP_IModuleHandler;
	ERRORHANDLER : L_IE1P_IErrorHandler;
	XSETERROR : BOOL;
	ESEVERITY : L_IE1P_SeverityLevel;
	WTEXTREFID : WORD;
	WERRORID : WORD;
	EREACTION : L_IE1P_Reaction;
	EGROUP : L_IE1P_Group;
	XERROR : BOOL;
	EERRORID : L_IE1P_Error;
	SCERRORINFORMATION : L_IE1P_ErrorInfo;
END_VAR
END_METHOD

METHOD SETREACTIONCOUNTERVARIABLE
VAR_INPUT
	EREACTIONNEW : L_IE1P_Reaction;
	DICOUNT : DINT;
END_VAR
VAR_IN_OUT
	REACTIONCOUNTER : L_IE1P_ReactionCounter;
END_VAR
END_METHOD

METHOD UPDATESEVERITYANDREACTIONCOUNTER
VAR_INPUT
	WMODE : WORD;
	ESEVERITYNEW : L_IE1P_SeverityLevel;
	EREACTIONNEW : L_IE1P_Reaction;
END_VAR
END_METHOD

METHOD FB_EXIT : BOOL
VAR_INPUT
	BINCOPYCODE : BOOL;
END_VAR
END_METHOD

METHOD FILLERRORATTRIBUTPARAMETER
VAR_INPUT
	ITFERRORATTRIBUTES : L_IE1P_IAttributes;
	IATTRIBUTNUMBER : INT;
END_VAR
VAR_IN_OUT
	PARAMETERITEM : L_IE1P_ParameterItemMid;
END_VAR
END_METHOD

METHOD FILLPLACEHODERPARAMETER
VAR_INPUT
	ITFTEXTPLACEHOLDER : L_IE1P_ITextPlaceHolder;
	PLACEHOLDERNBR : WORD;
END_VAR
VAR_IN_OUT
	PARAMINDEX : WORD;
	PARAMETERITEM : L_IE1P_ParameterItemMid;
END_VAR
END_METHOD

METHOD SENDERRORMSG
VAR_INPUT
	EGROUP : L_IE1P_Group;
END_VAR
END_METHOD

(* ---- L_IE1P_SETERRORSINGLESTRING.pou ---- *)
FUNCTION_BLOCK L_IE1P_SETERRORSINGLESTRING EXTENDS L_IE1P_SetErrorSingleBase
VAR_INPUT
	MODULEHANDLER : L_IMHP_IModuleHandler;
	ERRORHANDLER : L_IE1P_IErrorHandler;
	XSETERROR : BOOL;
	ESEVERITY : L_IE1P_SeverityLevel;
	WTEXTREFID : WORD;
	WERRORID : WORD;
	EREACTION : L_IE1P_Reaction := L_IE1P_Reaction.No_Reaction;
	EGROUP : L_IE1P_Group := L_IE1P_Group.ManufacturerGroup;
	STEXTPLACEHOLDER : STRING(50);
	ATTRIBUTES : L_IE1P_IAttributes;
END_VAR
VAR_OUTPUT
	XERROR : BOOL;
	EERRORID : L_IE1P_Error;
	SCERRORINFORMATION : L_IE1P_ErrorInfo;
END_VAR
VAR
	GETCONNECTEDMODULEHANDLER : L_IMHP_IModuleHandler;
	NBROFELEMENTS : WORD;
END_VAR
END_FUNCTION_BLOCK

METHOD GETPLACEHOLDERDATA : L_IE1P_PlaceHolderType
VAR_INPUT
	INDEX : WORD;
END_VAR
VAR_OUTPUT
	PDATA : POINTER TO BYTE;
END_VAR
END_METHOD

(* ---- L_IE1P_TEXTPLACEHOLDER.pou ---- *)
FUNCTION_BLOCK L_IE1P_TEXTPLACEHOLDER
VAR_INPUT
	EPLACEHOLDERTYPE1 : L_IE1P_PlaceHolderType;
	DIVALUE1 : DINT;
	DWVALUE1 : DWORD;
	SVALUE1 : STRING(50);
	EPLACEHOLDERTYPE2 : L_IE1P_PlaceHolderType;
	DIVALUE2 : DINT;
	DWVALUE2 : DWORD;
	SVALUE2 : STRING(50);
	EPLACEHOLDERTYPE3 : L_IE1P_PlaceHolderType;
	DIVALUE3 : DINT;
	DWVALUE3 : DWORD;
	SVALUE3 : STRING(50);
END_VAR
VAR
	NBROFELEMENTS : WORD;
END_VAR
END_FUNCTION_BLOCK

METHOD GETPLACEHOLDERDATA : L_IE1P_PlaceHolderType
VAR_INPUT
	INDEX : WORD;
END_VAR
VAR_OUTPUT
	PDATA : POINTER TO BYTE;
END_VAR
END_METHOD

(* ---- L_IE1P_TEXTPLACEHOLDERSINGLE.pou ---- *)
FUNCTION_BLOCK L_IE1P_TEXTPLACEHOLDERSINGLE
VAR_INPUT
	EPLACEHOLDERTYPE : L_IE1P_PlaceHolderType;
	DIVALUE : DINT;
	DWVALUE : DWORD;
	SVALUE : STRING(50);
END_VAR
VAR
	NBROFELEMENTS : WORD;
END_VAR
END_FUNCTION_BLOCK

METHOD GETPLACEHOLDERDATA : L_IE1P_PlaceHolderType
VAR_INPUT
	INDEX : WORD;
END_VAR
VAR_OUTPUT
	PDATA : POINTER TO BYTE;
END_VAR
END_METHOD
